(* IEC 61131-3 sources: PLC_ST_Simulator/examples/selftest, 4 files *)

(* ---- features.st ---- *)
TYPE E_Mode : (IDLE, RUN := 5, ERR); END_TYPE
TYPE ST_Pt : STRUCT x : INT := 3; y : REAL; END_STRUCT END_TYPE

VAR_GLOBAL
  gIn : BOOL;
  gCnt : INT;
  gArr : ARRAY[1..5] OF INT := [1, 2, 3(7)];
  gMode : E_Mode;
  gW : WORD := 16#00F0;
  gT : TIME;
END_VAR
VAR_GLOBAL CONSTANT
  N : INT := 5;
END_VAR

FUNCTION Add3 : INT
VAR_INPUT a, b : INT; c : INT := 100; END_VAR
Add3 := a + b + c;
END_FUNCTION

FUNCTION_BLOCK FB_Blink
VAR_INPUT en : BOOL; tOn : TIME := T#100ms; END_VAR
VAR_OUTPUT q : BOOL; END_VAR
VAR t1, t2 : TON; END_VAR
t1(IN := en AND NOT t2.Q, PT := tOn);
t2(IN := t1.Q, PT := tOn);
q := t1.Q;
END_FUNCTION_BLOCK

PROGRAM PLC_PRG
VAR
  i, sum : INT;
  overflow : INT := 32767;
  r : REAL;
  p : ST_Pt;
  blink : FB_Blink;
  ton1 : TON;
  ctu1 : CTU;
  rt : R_TRIG;
  s : STRING := 'abc';
  div : INT := 7;
  bits : BYTE;
  m2 : ARRAY[0..2, 0..1] OF DINT;
  res : INT;
END_VAR
sum := 0;
FOR i := 1 TO N DO
  IF i = 4 THEN CONTINUE; END_IF
  sum := sum + gArr[i];
END_FOR
overflow := overflow + 1;
r := INT_TO_REAL(div) / 2;
div := 7 / 2;
res := Add3(1, 2) + Add3(a := 1, b := 1, c := 1);
s := CONCAT(s, 'def');
bits := SHL(BYTE#1, 3) OR 2#1;
gW.0 := TRUE;
m2[2, 1] := 42;
gMode := E_Mode.RUN;
p.y := p.x * 1.5;
blink(en := gIn);
ton1(IN := gIn, PT := T#1s);
rt(CLK := gIn);
ctu1(CU := gIn, PV := 3);
IF rt.Q THEN gCnt := gCnt + 1; END_IF
gT := ton1.ET;
CASE gCnt OF
  0: ;
  1..2: i := 100;
ELSE
  i := -1;
END_CASE
WHILE i < 105 DO i := i + 1; IF i = 103 THEN EXIT; END_IF END_WHILE
END_PROGRAM

(* ---- konformitaet.st ---- *)
(* Konformität: Ganzzahl-Überlauf, Division, Bits, REAL, TIME, Strings, Kopiersemantik, Funktionen/FBs, Schleifen, CASE *)
TYPE ST_P : STRUCT x : INT; y : INT; a : ARRAY[0..2] OF INT; END_STRUCT END_TYPE
TYPE E_C : (ROT := 1, GRUEN := 2, BLAU := 4); END_TYPE

FUNCTION F_Out : INT
VAR_INPUT a : INT; END_VAR
VAR_OUTPUT doppelt : INT; END_VAR
VAR tmp : INT; END_VAR
tmp := tmp + 1;           (* Funktionen haben kein Gedächtnis *)
doppelt := a * 2;
F_Out := tmp;
END_FUNCTION

FUNCTION F_Early : INT
VAR_INPUT a : INT; END_VAR
F_Early := 1;
IF a > 0 THEN RETURN; END_IF
F_Early := 2;
END_FUNCTION

FUNCTION_BLOCK FB_Mem
VAR_INPUT inc : INT; END_VAR
VAR_OUTPUT sum : INT; END_VAR
VAR_TEMP t : INT; END_VAR
VAR n : INT; END_VAR
t := t + 1;      (* TEMP wird jedes Mal neu initialisiert *)
n := n + inc;
sum := n * 10 + t;
END_FUNCTION_BLOCK

FUNCTION_BLOCK FB_Swap
VAR_IN_OUT a, b : INT; END_VAR
VAR t : INT; END_VAR
t := a; a := b; b := t;
END_FUNCTION_BLOCK

PROGRAM PLC_PRG
VAR
    i : INT; si : SINT; usi : USINT; ui : UINT; di : DINT; ud : UDINT; li : LINT;
    b : BYTE; w : WORD; dw : DWORD;
    r : REAL; lr : LREAL;
    t : TIME;
    s : STRING; s5 : STRING(5);
    x : BOOL;
    p1, p2 : ST_P;
    a1, a2 : ARRAY[1..3] OF INT;
    m : ARRAY[1..2, 1..3] OF INT;
    c : E_C;
    fm : FB_Mem; fm2 : FB_Mem;
    sw : FB_Swap;
    o : INT; k : INT; n : INT;
END_VAR
;
END_PROGRAM

(* ---- oop.st ---- *)
(* Selbsttest: METHOD, ACTION, EXTENDS/SUPER^/THIS^, S=/R=, direkte Adressen, Pragmas *)
{attribute 'qualified_only'}
VAR_GLOBAL
    xTaster AT %IX0.0 : BOOL;
    xLampe  AT %QX0.0 : BOOL;
END_VAR

FUNCTION_BLOCK FB_Zaehler
VAR_INPUT  xEin : BOOL; END_VAR
VAR_OUTPUT iWert : INT; END_VAR
VAR rtEin : R_TRIG; END_VAR
rtEin(CLK := xEin);
IF rtEin.Q THEN Plus(n := 1); END_IF
END_FUNCTION_BLOCK

METHOD Plus : INT
VAR_INPUT n : INT; END_VAR
iWert := iWert + n;
Plus := iWert;
END_METHOD

ACTION Nullen:
iWert := 0;
END_ACTION

FUNCTION_BLOCK FB_Grenze EXTENDS FB_Zaehler
VAR_INPUT  iMax : INT := 3; END_VAR
VAR_OUTPUT xVoll : BOOL; END_VAR
SUPER^();
xVoll := THIS^.iWert >= iMax;
END_FUNCTION_BLOCK

PROGRAM PLC_PRG
VAR
    fb   : FB_Grenze;
    iRet : INT;
END_VAR
fb(xEin := %IX0.0);
IF fb.xVoll AND %IX0.1 THEN fb.Nullen(); END_IF
iRet := fb.Plus(n := 0);
xLampe S= fb.xVoll;
xLampe R= %IX0.1;
END_PROGRAM

(* ---- standard_fbs.st ---- *)
(* Standard-Bausteine: TON, TOF, TP, R_TRIG, F_TRIG, CTU, CTD, CTUD, SR, RS *)
PROGRAM PLC_PRG
VAR
    xIn : BOOL;
    ton1 : TON; tof1 : TOF; tp1 : TP;
    rt : R_TRIG; ft : F_TRIG;
    ctu1 : CTU; ctd1 : CTD; ctud1 : CTUD;
    sr1 : SR; rs1 : RS;
    xCu, xCd, xRes, xLoad, xS, xR : BOOL;
    nRt, nFt : INT;
END_VAR
ton1(IN := xIn, PT := T#100MS);
tof1(IN := xIn, PT := T#100MS);
tp1(IN := xIn, PT := T#100MS);
rt(CLK := xIn); IF rt.Q THEN nRt := nRt + 1; END_IF
ft(CLK := xIn); IF ft.Q THEN nFt := nFt + 1; END_IF
ctu1(CU := xCu, RESET := xRes, PV := 3);
ctd1(CD := xCd, LOAD := xLoad, PV := 2);
ctud1(CU := xCu, CD := xCd, RESET := xRes, LOAD := xLoad, PV := 2);
sr1(SET1 := xS, RESET := xR);
rs1(SET := xS, RESET1 := xR);
END_PROGRAM
